VAR_GLOBAL
    bFlag : BOOL;
    nCnt : DINT := 0; // cnt
END_VAR

(* stored: Version 1.1.0.1, ProductVersion 3.1.4026.18
   GVL GVL_Lint: Id {eeca5d67-1e2e-0cda-1cc0-d8d03086b510} *)
